Fanuc KAREL source: KO00073.KL

PROGRAM KO00073
%NOLOCKGROUP
%ENVIRONMENT MIR
VAR
  P1: XYZWPREXT
  P2: XYZWPREXT
  F: BOOLEAN
  OUT: POSITION
BEGIN
  F = TRUE
  OUT = MIRROR(P1, P2, F)
END KO00073
